(* IEC 61131-3 sources: volt/packages/volt-lsp-iec/test-corpus/twincat-project14/TwinCAT Project14/PLC/Untitled2/Untitled2 Project/References/Tc2_System, 164 files *)

(* ---- E_AdsErr.dut ---- *)
TYPE E_AdsErr :
(
	NOERR,
	ROUTER_NOLOCKEDMEMORY,
	ROUTER_RESIZEMEMORY,
	ROUTER_MAILBOXFULL,
	ROUTER_DEBUGBOXFULL,
	ROUTER_UNKNOWNPORTTYPE,
	ROUTER_NOTINITIALIZED,
	ROUTER_PORTALREADYINUSE,
	ROUTER_NOTREGISTERED,
	ROUTER_NOMOREQUEUES,
	ROUTER_INVALIDPORT,
	ROUTER_NOTACTIVATED,
	ROUTER_FRAGMENTBOXFULL,
	ROUTER_FRAGMENTTIMEOUT,
	ROUTER_TOBEREMOVED,
	DEVICE_ERROR,
	DEVICE_SRVNOTSUPP,
	DEVICE_INVALIDGRP,
	DEVICE_INVALIDOFFSET,
	DEVICE_INVALIDACCESS,
	DEVICE_INVALIDSIZE,
	DEVICE_INVALIDDATA,
	DEVICE_NOTREADY,
	DEVICE_BUSY,
	DEVICE_INVALIDCONTEXT,
	DEVICE_NOMEMORY,
	DEVICE_INVALIDPARM,
	DEVICE_NOTFOUND,
	DEVICE_SYNTAX,
	DEVICE_INCOMPATIBLE,
	DEVICE_EXISTS,
	DEVICE_SYMBOLNOTFOUND,
	DEVICE_SYMBOLVERSIONINVALID,
	DEVICE_INVALIDSTATE,
	DEVICE_TRANSMODENOTSUPP,
	DEVICE_NOTIFYHNDINVALID,
	DEVICE_CLIENTUNKNOWN,
	DEVICE_NOMOREHDLS,
	DEVICE_INVALIDWATCHSIZE,
	DEVICE_NOTINIT,
	DEVICE_TIMEOUT,
	DEVICE_NOINTERFACE,
	DEVICE_INVALIDINTERFACE,
	DEVICE_INVALIDCLSID,
	DEVICE_INVALIDOBJID,
	DEVICE_PENDING,
	DEVICE_ABORTED,
	DEVICE_WARNING,
	DEVICE_INVALIDARRAYIDX,
	DEVICE_SYMBOLNOTACTIVE,
	DEVICE_ACCESSDENIED,
	DEVICE_LICENSENOTFOUND,
	DEVICE_LICENSEEXPIRED,
	DEVICE_LICENSEEXCEEDED,
	DEVICE_LICENSEINVALID,
	DEVICE_LICENSESYSTEMID,
	DEVICE_LICENSENOTIMELIMIT,
	DEVICE_LICENSEFUTUREISSUE,
	DEVICE_LICENSETIMETOLONG,
	DEVICE_EXCEPTION,
	DEVICE_LICENSEDUPLICATED,
	CLIENT_ERROR,
	CLIENT_INVALIDPARM,
	CLIENT_LISTEMPTY,
	CLIENT_VARUSED,
	CLIENT_DUPLINVOKEID,
	CLIENT_SYNCTIMEOUT,
	CLIENT_W32ERROR,
	CLIENT_TIMEOUTINVALID,
	CLIENT_PORTNOTOPEN,
	CLIENT_NOAMSADDR,
	CLIENT_SYNCINTERNAL,
	CLIENT_ADDHASH,
	CLIENT_REMOVEHASH,
	CLIENT_NOMORESYM,
	CLIENT_SYNCRESINVALID,
	CLIENT_SYNCPORTLOCKED
);
END_TYPE

(* ---- E_HRESULTAdsErr.dut ---- *)
TYPE E_HRESULTAdsErr :
(
	HRESULT_ADS_NOERROR,
	ROUTER_NOLOCKEDMEMORY,
	ROUTER_RESIZEMEMORY,
	ROUTER_MAILBOXFULL,
	ROUTER_DEBUGBOXFULL,
	ROUTER_UNKNOWNPORTTYPE,
	ROUTER_NOTINITIALIZED,
	ROUTER_PORTALREADYINUSE,
	ROUTER_NOTREGISTERED,
	ROUTER_NOMOREQUEUES,
	ROUTER_INVALIDPORT,
	ROUTER_NOTACTIVATED,
	ROUTER_FRAGMENTBOXFULL,
	ROUTER_FRAGMENTTIMEOUT,
	ROUTER_TOBEREMOVED,
	ERROR,
	SRVNOTSUPP,
	INVALIDGRP,
	INVALIDOFFSET,
	INVALIDACCESS,
	INVALIDSIZE,
	INVALIDDATA,
	NOTREADY,
	BUSY,
	INVALIDCONTEXT,
	NOMEMORY,
	INVALIDPARM,
	NOTFOUND,
	SYNTAX,
	INCOMPATIBLE,
	EXISTS,
	SYMBOLNOTFOUND,
	SYMBOLVERSIONINVALID,
	INVALIDSTATE,
	TRANSMODENOTSUPP,
	NOTIFYHNDINVALID,
	CLIENTUNKNOWN,
	NOMOREHDLS,
	INVALIDWATCHSIZE,
	NOTINIT,
	TIMEOUT,
	NOINTERFACE,
	INVALIDINTERFACE,
	INVALIDCLSID,
	INVALIDOBJID,
	PENDING,
	ABORTED,
	WARNING,
	INVALIDARRAYIDX,
	SYMBOLNOTACTIVE,
	ACCESSDENIED,
	LICENSENOTFOUND,
	LICENSEEXPIRED,
	LICENSEEXCEEDED,
	LICENSEINVALID,
	LICENSESYSTEMID,
	LICENSENOTIMELIMIT,
	LICENSEFUTUREISSUE,
	LICENSETIMETOLONG,
	EXCEPTION,
	LICENSEDUPLICATED,
	CLIENT_ERROR,
	CLIENT_INVALIDPARM,
	CLIENT_LISTEMPTY,
	CLIENT_VARUSED,
	CLIENT_DUPLINVOKEID,
	CLIENT_SYNCTIMEOUT,
	CLIENT_W32ERROR,
	CLIENT_TIMEOUTINVALID,
	CLIENT_PORTNOTOPEN,
	CLIENT_NOAMSADDR,
	CLIENT_SYNCINTERNAL,
	CLIENT_ADDHASH,
	CLIENT_REMOVEHASH,
	CLIENT_NOMORESYM,
	CLIENT_SYNCRESINVALID,
	CLIENT_SYNCPORTLOCKED
);
END_TYPE

(* ---- E_OpenPath.dut ---- *)
TYPE E_OpenPath :
(
	PATH_GENERIC,
	PATH_BOOTPRJ,
	PATH_BOOTDATA,
	PATH_BOOTPATH,
	PATH_USERPATH1,
	PATH_USERPATH2,
	PATH_USERPATH3,
	PATH_USERPATH4,
	PATH_USERPATH5,
	PATH_USERPATH6,
	PATH_USERPATH7,
	PATH_USERPATH8,
	PATH_USERPATH9
);
END_TYPE

(* ---- E_SeekOrigin.dut ---- *)
TYPE E_SeekOrigin :
(
	SEEK_SET,
	SEEK_CUR,
	SEEK_END
);
END_TYPE

(* ---- E_TcEventClass.dut ---- *)
TYPE E_TcEventClass :
(
	TCEVENTCLASS_NONE,
	TCEVENTCLASS_MAINTENANCE,
	TCEVENTCLASS_MESSAGE,
	TCEVENTCLASS_HINT,
	TCEVENTCLASS_STATEINFO,
	TCEVENTCLASS_INSTRUCTION,
	TCEVENTCLASS_WARNING,
	TCEVENTCLASS_ALARM,
	TCEVENTCLASS_PARAMERROR
);
END_TYPE

(* ---- E_TcEventClearModes.dut ---- *)
TYPE E_TcEventClearModes :
(
	TCEVENTLOGIOFFS_CLEARACTIVE,
	TCEVENTLOGIOFFS_CLEARLOGGED,
	TCEVENTLOGIOFFS_CLEARALL
);
END_TYPE

(* ---- E_TcEventPriority.dut ---- *)
TYPE E_TcEventPriority :
(
	TCEVENTPRIO_IMPLICIT
);
END_TYPE

(* ---- E_TcEventStreamType.dut ---- *)
TYPE E_TcEventStreamType :
(
	TCEVENTSTREAM_INVALID,
	TCEVENTSTREAM_SIMPLE,
	TCEVENTSTREAM_NORMAL,
	TCEVENTSTREAM_NOSOURCE,
	TCEVENTSTREAM_CLASSID,
	TCEVENTSTREAM_CLSNOSRC,
	TCEVENTSTREAM_READCLASSCOUNT,
	TCEVENTSTREAM_MAXTYPE
);
END_TYPE

(* ---- E_TcMemoryArea.dut ---- *)
TYPE E_TcMemoryArea :
(
	Unknown,
	Static,
	Dynamic,
	CNC
);
END_TYPE

(* ---- E_UsrLED_Color.dut ---- *)
TYPE E_UsrLED_Color :
(
	eUsrLED_Off,
	eUsrLED_Red,
	eUsrLED_Blue,
	eUsrLED_Green
);
END_TYPE

(* ---- E_WATCHDOG_TIME_CONFIG.dut ---- *)
TYPE E_WATCHDOG_TIME_CONFIG :
(
	eWATCHDOG_TIME_DISABLED,
	eWATCHDOG_TIME_SECONDS,
	eWATCHDOG_TIME_MINUTES
);
END_TYPE

(* ---- FW_NoOfByte.dut ---- *)
TYPE FW_NoOfByte :
(
	NoOfByte_Byte,
	NoOfByte_Word,
	NoOfByte_DWord
);
END_TYPE

(* ---- Global_Variables.gvl ---- *)
VAR_GLOBAL
	AMSPORT_LOGGER : UINT;
	AMSPORT_EVENTLOG : UINT;
	AMSPORT_R0_RTIME : UINT;
	AMSPORT_R0_IO : UINT;
	AMSPORT_R0_NC : UINT;
	AMSPORT_R0_NCSAF : UINT;
	AMSPORT_R0_NCSVB : UINT;
	AMSPORT_R0_ISG : UINT;
	AMSPORT_R0_CNC : UINT;
	AMSPORT_R0_LINE : UINT;
	AMSPORT_R0_PLC : UINT;
	AMSPORT_R0_PLC_RTS1 : UINT;
	AMSPORT_R0_PLC_RTS2 : UINT;
	AMSPORT_R0_PLC_RTS3 : UINT;
	AMSPORT_R0_PLC_RTS4 : UINT;
	AMSPORT_R0_CAM : UINT;
	AMSPORT_R0_CAMTOOL : UINT;
	AMSPORT_R3_SYSSERV : UINT;
	AMSPORT_R3_SCOPESERVER : UINT;
	ADSSTATE_INVALID : UINT;
	ADSSTATE_IDLE : UINT;
	ADSSTATE_RESET : UINT;
	ADSSTATE_INIT : UINT;
	ADSSTATE_START : UINT;
	ADSSTATE_RUN : UINT;
	ADSSTATE_STOP : UINT;
	ADSSTATE_SAVECFG : UINT;
	ADSSTATE_LOADCFG : UINT;
	ADSSTATE_POWERFAILURE : UINT;
	ADSSTATE_POWERGOOD : UINT;
	ADSSTATE_ERROR : UINT;
	ADSSTATE_SHUTDOWN : UINT;
	ADSSTATE_SUSPEND : UINT;
	ADSSTATE_RESUME : UINT;
	ADSSTATE_CONFIG : UINT;
	ADSSTATE_RECONFIG : UINT;
	ADSSTATE_STOPPING : UINT;
	ADSSTATE_INCOMPATIBLE : UINT;
	ADSSTATE_EXCEPTION : UINT;
	ADSSTATE_MAXSTATES : UINT;
	ADSIGRP_SYMTAB : UDINT;
	ADSIGRP_SYMNAME : UDINT;
	ADSIGRP_SYMVAL : UDINT;
	ADSIGRP_SYM_HNDBYNAME : UDINT;
	ADSIGRP_SYM_VALBYNAME : UDINT;
	ADSIGRP_SYM_VALBYHND : UDINT;
	ADSIGRP_SYM_RELEASEHND : UDINT;
	ADSIGRP_SYM_INFOBYNAME : UDINT;
	ADSIGRP_SYM_VERSION : UDINT;
	ADSIGRP_SYM_INFOBYNAMEEX : UDINT;
	ADSIGRP_SYM_DOWNLOAD : UDINT;
	ADSIGRP_SYM_UPLOAD : UDINT;
	ADSIGRP_SYM_UPLOADINFO : UDINT;
	ADSIGRP_SYMNOTE : UDINT;
	ADSIGRP_IOIMAGE_RWIB : UDINT;
	ADSIGRP_IOIMAGE_RWIX : UDINT;
	ADSIGRP_IOIMAGE_RISIZE : UDINT;
	ADSIGRP_IOIMAGE_RWOB : UDINT;
	ADSIGRP_IOIMAGE_RWOX : UDINT;
	ADSIGRP_IOIMAGE_ROSIZE : UDINT;
	ADSIGRP_IOIMAGE_CLEARI : UDINT;
	ADSIGRP_IOIMAGE_CLEARO : UDINT;
	ADSIGRP_IOIMAGE_RWIOB : UDINT;
	ADSIGRP_DEVICE_DATA : UDINT;
	ADSIOFFS_DEVDATA_ADSSTATE : UDINT;
	ADSIOFFS_DEVDATA_DEVSTATE : UDINT;
	SYSTEMSERVICE_OPENCREATE : UDINT;
	SYSTEMSERVICE_OPENREAD : UDINT;
	SYSTEMSERVICE_OPENWRITE : UDINT;
	SYSTEMSERVICE_CREATEFILE : UDINT;
	SYSTEMSERVICE_CLOSEHANDLE : UDINT;
	SYSTEMSERVICE_FOPEN : UDINT;
	SYSTEMSERVICE_FCLOSE : UDINT;
	SYSTEMSERVICE_FREAD : UDINT;
	SYSTEMSERVICE_FWRITE : UDINT;
	SYSTEMSERVICE_FSEEK : UDINT;
	SYSTEMSERVICE_FTELL : UDINT;
	SYSTEMSERVICE_FGETS : UDINT;
	SYSTEMSERVICE_FPUTS : UDINT;
	SYSTEMSERVICE_FSCANF : UDINT;
	SYSTEMSERVICE_FPRINTF : UDINT;
	SYSTEMSERVICE_FEOF : UDINT;
	SYSTEMSERVICE_FDELETE : UDINT;
	SYSTEMSERVICE_FRENAME : UDINT;
	SYSTEMSERVICE_MKDIR : UDINT;
	SYSTEMSERVICE_RMDIR : UDINT;
	SYSTEMSERVICE_REG_HKEYLOCALMACHINE : UDINT;
	SYSTEMSERVICE_SENDEMAIL : UDINT;
	SYSTEMSERVICE_TIMESERVICES : UDINT;
	SYSTEMSERVICE_STARTPROCESS : UDINT;
	SYSTEMSERVICE_CHANGENETID : UDINT;
	TIMESERVICE_DATEANDTIME : UDINT;
	TIMESERVICE_SYSTEMTIMES : UDINT;
	TIMESERVICE_RTCTIMEDIFF : UDINT;
	TIMESERVICE_ADJUSTTIMETORTC : UDINT;
	TIMESERVICE_TIMEZONINFORMATION : UDINT;
	ADSLOG_MSGTYPE_HINT : DWORD;
	ADSLOG_MSGTYPE_WARN : DWORD;
	ADSLOG_MSGTYPE_ERROR : DWORD;
	ADSLOG_MSGTYPE_LOG : DWORD;
	ADSLOG_MSGTYPE_MSGBOX : DWORD;
	ADSLOG_MSGTYPE_RESOURCE : DWORD;
	ADSLOG_MSGTYPE_STRING : DWORD;
	BOOTDATAFLAGS_RETAIN_LOADED : BYTE;
	BOOTDATAFLAGS_RETAIN_INVALID : BYTE;
	BOOTDATAFLAGS_RETAIN_REQUESTED : BYTE;
	BOOTDATAFLAGS_PERSISTENT_LOADED : BYTE;
	BOOTDATAFLAGS_PERSISTENT_INVALID : BYTE;
	SYSTEMSTATEFLAGS_BSOD : BYTE;
	SYSTEMSTATEFLAGS_RTVIOLATION : BYTE;
	FOPEN_MODEREAD : DWORD;
	FOPEN_MODEWRITE : DWORD;
	FOPEN_MODEAPPEND : DWORD;
	FOPEN_MODEPLUS : DWORD;
	FOPEN_MODEBINARY : DWORD;
	FOPEN_MODETEXT : DWORD;
	FILE_OPENCREATE : DWORD;
	FILE_OPENREAD : DWORD;
	FILE_OPENWRITE : DWORD;
	FILE_READ : DWORD;
	FILE_WRITE : DWORD;
	FILE_SEEKBEGIN : DWORD;
	FILE_SEEKEND : DWORD;
	TCEVENTFLAG_PRIOCLASS : WORD;
	TCEVENTFLAG_FMTSELF : WORD;
	TCEVENTFLAG_LOG : WORD;
	TCEVENTFLAG_MSGBOX : WORD;
	TCEVENTFLAG_SRCID : WORD;
	TCEVENTFLAG_AUTOFMTALL : WORD;
	TCEVENTSTATE_INVALID : WORD;
	TCEVENTSTATE_SIGNALED : WORD;
	TCEVENTSTATE_RESET : WORD;
	TCEVENTSTATE_CONFIRMED : WORD;
	TCEVENTSTATE_RESETCON : WORD;
	TCEVENT_SRCNAMESIZE : INT;
	TCEVENT_FMTPRGSIZE : INT;
	PI : LREAL;
	DEFAULT_ADS_TIMEOUT : TIME;
	MAX_STRING_LENGTH : UDINT;
	MAX_TCBADEV_USERDATA : UDINT;
	SYSTEMSERVICE_BADEVAPI : UDINT;
	BADEVAPIIGRP_GENERAL : UDINT;
	BADEVAPIIOFFS_GENERAL_VERSION : UDINT;
	BIOSIGRP_WATCHDOG : UDINT;
	BIOSIOFFS_WATCHDOG_ENABLE : UDINT;
	BIOSIOFFS_WATCHDOG_CONFIG : UDINT;
	BIOSIOFFS_WATCHDOG_GET_WD_CONFIG : UDINT;
	BIOSIOFFS_WATCHDOG_SET_WD_CONFIG : UDINT;
	BIOSIOFFS_WATCHDOG_ACTIVATE_PWCTR_IO : UDINT;
	BIOSIOFFS_WATCHDOG_TRIG_WD_TIMESPAN : UDINT;
	BIOSIOFFS_WATCHDOG_IO_RETRIGGER : UDINT;
	BIOSIOFFS_WATCHDOG_GET_IO_ADDR : UDINT;
	BIOSIOFFS_WATCHDOG_GET_IO_ADDR_EX : UDINT;
	BIOSIGRP_LED : UDINT;
	BIOSIOFFS_LED_SET_USER : UDINT;
	BIOSIOFFS_LED_SET_USER2 : UDINT;
END_VAR

(* ---- Global_Version.gvl ---- *)
VAR_GLOBAL
	stLibVersion_Tc2_System : ST_LibVersion;
END_VAR

(* ---- Param.gvl ---- *)
VAR_GLOBAL
	TABLE_UPPER_BOUND : INT;
	STRING_LENGTH_EXP : INT;
	STRING_LENGTH_ADDRESS : INT;
	STRING_LENGTH_COMMENT : INT;
	STRING_LENGTH_OUTSTRING : INT;
	TABLE_SHOW_VALID_ITEMS : BOOL;
END_VAR

(* ---- AdsErr_TO_HRESULTAdsErr.pou ---- *)
FUNCTION AdsErr_TO_HRESULTAdsErr : E_HRESULTAdsErr
VAR_INPUT
	eErrId : E_AdsErr;
END_VAR
END_FUNCTION

(* ---- ADSLOGDINT.pou ---- *)
FUNCTION ADSLOGDINT : DINT
VAR_INPUT
	msgCtrlMask : DWORD;
	msgFmtStr : T_MaxString;
	dintArg : DINT;
END_VAR
END_FUNCTION

(* ---- ADSLOGLREAL.pou ---- *)
FUNCTION ADSLOGLREAL : DINT
VAR_INPUT
	msgCtrlMask : DWORD;
	msgFmtStr : T_MaxString;
	lrealArg : LREAL;
END_VAR
END_FUNCTION

(* ---- ADSLOGSTR.pou ---- *)
FUNCTION ADSLOGSTR : DINT
VAR_INPUT
	msgCtrlMask : DWORD;
	msgFmtStr : T_MaxString;
	strArg : T_MaxString;
END_VAR
END_FUNCTION

(* ---- AppendErrorString.pou ---- *)
FUNCTION AppendErrorString
VAR_IN_OUT
	strOld : STRING(STRING_LENGTH_EXP);
	strNew : STRING(1);
END_VAR
END_FUNCTION

(* ---- BAVERSION_TO_DWORD.pou ---- *)
FUNCTION BAVERSION_TO_DWORD : DWORD
VAR_INPUT
	nVersion : BYTE;
	nRevision : BYTE;
	nBuild : WORD;
END_VAR
END_FUNCTION

(* ---- CLEARBIT32.pou ---- *)
FUNCTION CLEARBIT32 : DWORD
VAR_INPUT
	inVal32 : DWORD;
	bitNo : SINT;
END_VAR
END_FUNCTION

(* ---- CONCATX.pou ---- *)
FUNCTION CONCATX
VAR_IN_OUT
	STR1 : STRING(STRING_LENGTH_EXP);
	STR2 : STRING(1);
END_VAR
END_FUNCTION

(* ---- CSETBIT32.pou ---- *)
FUNCTION CSETBIT32 : DWORD
VAR_INPUT
	inVal32 : DWORD;
	bitNo : SINT;
	bitVal : BOOL;
END_VAR
END_FUNCTION

(* ---- F_CheckMemoryArea.pou ---- *)
FUNCTION F_CheckMemoryArea : E_TcMemoryArea
VAR_INPUT
	pData : PVOID;
	nSize : UDINT;
END_VAR
END_FUNCTION

(* ---- F_CmpLibVersion.pou ---- *)
FUNCTION F_CmpLibVersion : DINT
VAR_INPUT
	stVersion : ST_LibVersion;
	iMajor : UINT;
	iMinor : UINT;
	iBuild : UINT;
	iRevision : UINT;
END_VAR
END_FUNCTION

(* ---- F_CompareFwVersion.pou ---- *)
FUNCTION F_CompareFwVersion : BOOL
VAR_INPUT
	major : UINT;
	minor : UINT;
	revision : UINT;
	patch : UINT;
END_VAR
END_FUNCTION

(* ---- F_CreateAmsNetId.pou ---- *)
FUNCTION F_CreateAmsNetId : T_AmsNetId
VAR_INPUT
	nIds : T_AmsNetIdArr;
END_VAR
END_FUNCTION

(* ---- F_CreateIPv4Addr.pou ---- *)
FUNCTION F_CreateIPv4Addr : T_IPv4Addr
VAR_INPUT
	nIds : T_IPv4AddrArr;
END_VAR
END_FUNCTION

(* ---- F_CreateMacAddr.pou ---- *)
FUNCTION F_CreateMacAddr : T_MacAddr
VAR_INPUT
	aMacAddr : T_MacAddrArr;
	sSeparator : STRING(1);
	bLoCase : BOOL;
END_VAR
END_FUNCTION

(* ---- F_GetCpuCoreIndex.pou ---- *)
FUNCTION F_GetCpuCoreIndex : DINT
VAR_INPUT
	nTaskIndex : DINT;
END_VAR
END_FUNCTION

(* ---- F_GetCpuCoreInfo.pou ---- *)
FUNCTION F_GetCpuCoreInfo : HRESULT
VAR_INPUT
	nCpuCoreIndex : DINT;
	pInfo : POINTER TO ST_CpuCoreInfo;
END_VAR
END_FUNCTION

(* ---- F_GetMappingPartner.pou ---- *)
FUNCTION F_GetMappingPartner : OTCID
VAR_INPUT
	p : PVOID;
	n : UDINT;
END_VAR
END_FUNCTION

(* ---- F_GetMappingStatus.pou ---- *)
FUNCTION F_GetMappingStatus : EPlcMappingStatus
VAR_INPUT
	p : PVOID;
	n : UDINT;
END_VAR
END_FUNCTION

(* ---- F_GetStructMemberAlignment.pou ---- *)
FUNCTION F_GetStructMemberAlignment : BYTE
END_FUNCTION

(* ---- F_GetSystemTime.pou ---- *)
FUNCTION F_GetSystemTime : ULINT
END_FUNCTION

(* ---- F_GetTaskInfo.pou ---- *)
FUNCTION F_GetTaskInfo : PlcTaskSystemInfo
END_FUNCTION

(* ---- F_GetTaskTime.pou ---- *)
FUNCTION F_GetTaskTime : ULINT
END_FUNCTION

(* ---- F_GetTaskTotalTime.pou ---- *)
FUNCTION F_GetTaskTotalTime : UDINT
VAR_INPUT
	nTaskIndex : DINT;
END_VAR
END_FUNCTION

(* ---- F_GetVersionTcSystem.pou ---- *)
FUNCTION F_GetVersionTcSystem : UINT
VAR_INPUT
	nVersionElement : INT;
END_VAR
END_FUNCTION

(* ---- F_IOPortRead.pou ---- *)
FUNCTION F_IOPortRead : DWORD
VAR_INPUT
	nAddr : UDINT;
	eSize : E_IOAccessSize;
END_VAR
END_FUNCTION

(* ---- F_IOPortWrite.pou ---- *)
FUNCTION F_IOPortWrite : BOOL
VAR_INPUT
	nAddr : UDINT;
	eSize : E_IOAccessSize;
	nValue : DWORD;
END_VAR
END_FUNCTION

(* ---- F_RaiseException.pou ---- *)
FUNCTION F_RaiseException
VAR_INPUT
	exceptionCode : UDINT;
END_VAR
END_FUNCTION

(* ---- F_ScanAmsNetIds.pou ---- *)
FUNCTION F_ScanAmsNetIds : T_AmsNetIdArr
VAR_INPUT
	sNetID : T_AmsNetID;
END_VAR
END_FUNCTION

(* ---- F_ScanIPv4AddrIds.pou ---- *)
FUNCTION F_ScanIPv4AddrIds : T_IPv4AddrArr
VAR_INPUT
	sIPv4 : T_IPv4Addr;
END_VAR
END_FUNCTION

(* ---- F_SplitPathName.pou ---- *)
FUNCTION F_SplitPathName : BOOL
VAR_INPUT
	sPathName : T_MaxString;
END_VAR
VAR_IN_OUT
	sDrive : STRING(3);
	sDir : T_MaxString;
	sFileName : T_MaxString;
	sExt : T_MaxString;
END_VAR
END_FUNCTION

(* ---- F_ToASC.pou ---- *)
FUNCTION F_ToASC : BYTE
VAR_INPUT
	str : STRING;
END_VAR
END_FUNCTION

(* ---- F_ToCHR.pou ---- *)
FUNCTION F_ToCHR : STRING
VAR_INPUT
	c : BYTE;
END_VAR
END_FUNCTION

(* ---- FW_AdsLogDINT.pou ---- *)
FUNCTION FW_AdsLogDINT : DINT
VAR_INPUT
	nCtrlMask : DWORD;
	sMsgFmt : STRING(255);
	nArg : DINT;
END_VAR
END_FUNCTION

(* ---- FW_AdsLogLREAL.pou ---- *)
FUNCTION FW_AdsLogLREAL : DINT
VAR_INPUT
	nCtrlMask : DWORD;
	sMsgFmt : STRING(255);
	fArg : LREAL;
END_VAR
END_FUNCTION

(* ---- FW_AdsLogSTR.pou ---- *)
FUNCTION FW_AdsLogSTR : DINT
VAR_INPUT
	nCtrlMask : DWORD;
	sMsgFmt : STRING(255);
	sArg : STRING(255);
END_VAR
END_FUNCTION

(* ---- FW_GetCpuIndex.pou ---- *)
FUNCTION FW_GetCpuIndex : DINT
VAR_INPUT
	taskIndex : DINT;
END_VAR
END_FUNCTION

(* ---- FW_GetCpuInfo.pou ---- *)
FUNCTION FW_GetCpuInfo : HRESULT
VAR_INPUT
	cpuIndex : DINT;
	pInfo : POINTER TO ST_CpuCoreInfo;
END_VAR
END_FUNCTION

(* ---- FW_GetCurTaskIndexEx.pou ---- *)
FUNCTION FW_GetCurTaskIndexEx : DINT
END_FUNCTION

(* ---- FW_GetMappingPartner.pou ---- *)
FUNCTION FW_GetMappingPartner : OTCID
VAR_INPUT
	p : PVOID;
	n : UDINT;
END_VAR
END_FUNCTION

(* ---- FW_GetMappingStatus.pou ---- *)
FUNCTION FW_GetMappingStatus : EPlcMappingStatus
VAR_INPUT
	p : PVOID;
	n : UDINT;
END_VAR
END_FUNCTION

(* ---- FW_GetTaskTotalTime.pou ---- *)
FUNCTION FW_GetTaskTotalTime : UDINT
VAR_INPUT
	taskIndex : DINT;
END_VAR
END_FUNCTION

(* ---- FW_GetVersionTcBase.pou ---- *)
FUNCTION FW_GetVersionTcBase : UINT
VAR_INPUT
	nVersionElement : INT;
END_VAR
END_FUNCTION

(* ---- FW_LptSignal.pou ---- *)
FUNCTION FW_LptSignal : BOOL
VAR_INPUT
	nPortAddr : UINT;
	nPinNo : UINT;
	bOnOff : BOOL;
END_VAR
END_FUNCTION

(* ---- FW_MemCmp.pou ---- *)
FUNCTION FW_MemCmp : DINT
VAR_INPUT
	pBuf1 : PVOID;
	pBuf2 : PVOID;
	cbLen : UDINT;
END_VAR
END_FUNCTION

(* ---- FW_MemCpy.pou ---- *)
FUNCTION FW_MemCpy : UDINT
VAR_INPUT
	pDest : PVOID;
	pSrc : PVOID;
	cbLen : UDINT;
END_VAR
END_FUNCTION

(* ---- FW_MemMove.pou ---- *)
FUNCTION FW_MemMove : UDINT
VAR_INPUT
	pDest : PVOID;
	pSrc : PVOID;
	cbLen : UDINT;
END_VAR
END_FUNCTION

(* ---- FW_MemSet.pou ---- *)
FUNCTION FW_MemSet : UDINT
VAR_INPUT
	pDest : PVOID;
	nFillByte : USINT;
	cbLen : UDINT;
END_VAR
END_FUNCTION

(* ---- FW_PortRead.pou ---- *)
FUNCTION FW_PortRead : DWORD
VAR_INPUT
	nPortAddr : UDINT;
	eNoOfByte : FW_NoOfByte;
END_VAR
END_FUNCTION

(* ---- FW_PortWrite.pou ---- *)
FUNCTION FW_PortWrite : BOOL
VAR_INPUT
	nPortAddr : UDINT;
	eNoOfByte : FW_NoOfByte;
	nValue : DWORD;
END_VAR
END_FUNCTION

(* ---- FW_RaiseException.pou ---- *)
FUNCTION FW_RaiseException
VAR_INPUT
	exceptionCode : UDINT;
END_VAR
END_FUNCTION

(* ---- GETBIT32.pou ---- *)
FUNCTION GETBIT32 : BOOL
VAR_INPUT
	inVal32 : DWORD;
	bitNo : SINT;
END_VAR
END_FUNCTION

(* ---- GETCURTASKINDEXEX.pou ---- *)
FUNCTION GETCURTASKINDEXEX : DINT
END_FUNCTION

(* ---- HRESULTAdsErr_TO_AdsErr.pou ---- *)
FUNCTION HRESULTAdsErr_TO_AdsErr : E_AdsErr
VAR_INPUT
	hrErrId : E_HRESULTAdsErr;
END_VAR
END_FUNCTION

(* ---- LPTSIGNAL.pou ---- *)
FUNCTION LPTSIGNAL : BOOL
VAR_INPUT
	PortAddr : UINT;
	PinNo : UINT;
	OnOff : BOOL;
END_VAR
END_FUNCTION

(* ---- MEMCMP.pou ---- *)
FUNCTION MEMCMP : DINT
VAR_INPUT
	pBuf1 : PVOID;
	pBuf2 : PVOID;
	n : UDINT;
END_VAR
END_FUNCTION

(* ---- MEMCPY.pou ---- *)
FUNCTION MEMCPY : UDINT
VAR_INPUT
	destAddr : PVOID;
	srcAddr : PVOID;
	n : UDINT;
END_VAR
END_FUNCTION

(* ---- MEMMOVE.pou ---- *)
FUNCTION MEMMOVE : UDINT
VAR_INPUT
	destAddr : PVOID;
	srcAddr : PVOID;
	n : UDINT;
END_VAR
END_FUNCTION

(* ---- MEMSET.pou ---- *)
FUNCTION MEMSET : UDINT
VAR_INPUT
	destAddr : PVOID;
	fillByte : USINT;
	n : UDINT;
END_VAR
END_FUNCTION

(* ---- ROL32.pou ---- *)
FUNCTION ROL32 : DWORD
VAR_INPUT
	inVal32 : DWORD;
	n : SINT;
END_VAR
END_FUNCTION

(* ---- ROR32.pou ---- *)
FUNCTION ROR32 : DWORD
VAR_INPUT
	inVal32 : DWORD;
	n : SINT;
END_VAR
END_FUNCTION

(* ---- SETBIT32.pou ---- *)
FUNCTION SETBIT32 : DWORD
VAR_INPUT
	inVal32 : DWORD;
	bitNo : SINT;
END_VAR
END_FUNCTION

(* ---- SHL32.pou ---- *)
FUNCTION SHL32 : DWORD
VAR_INPUT
	inVal32 : DWORD;
	n : SINT;
END_VAR
END_FUNCTION

(* ---- SHR32.pou ---- *)
FUNCTION SHR32 : DWORD
VAR_INPUT
	inVal32 : DWORD;
	n : SINT;
END_VAR
END_FUNCTION

(* ---- TestAndSet.pou ---- *)
FUNCTION TestAndSet : BOOL
VAR_IN_OUT
	Flag : BOOL;
END_VAR
END_FUNCTION

(* ---- ADSCLEAREVENTS.pou ---- *)
FUNCTION_BLOCK ADSCLEAREVENTS
VAR_INPUT
	NetID : T_AmsNetId;
	bClear : BOOL;
	iMode : UDINT;
	tTimeout : TIME;
END_VAR
VAR_OUTPUT
	bBusy : BOOL;
	bErr : BOOL;
	iErrId : UDINT;
END_VAR
END_FUNCTION_BLOCK

(* ---- ADSLOGEVENT.pou ---- *)
FUNCTION_BLOCK ADSLOGEVENT
VAR_INPUT
	NETID : T_AmsNetId;
	PORT : UINT;
	Event : BOOL;
	EventQuit : BOOL;
	EventConfigData : TcEvent;
	EventDataAddress : PVOID;
	EventDataLength : UDINT;
	FbCleanup : BOOL;
	TMOUT : TIME;
END_VAR
VAR_OUTPUT
	EventState : UDINT;
	Err : BOOL;
	ErrId : UDINT;
	Quit : BOOL;
END_VAR
END_FUNCTION_BLOCK

(* ---- ADSRDDEVINFO.pou ---- *)
FUNCTION_BLOCK ADSRDDEVINFO
VAR_INPUT
	NETID : T_AmsNetId;
	PORT : T_AmsPort;
	RDINFO : BOOL;
	TMOUT : TIME;
END_VAR
VAR_OUTPUT
	BUSY : BOOL;
	ERR : BOOL;
	ERRID : UDINT;
	DEVNAME : STRING(19);
	DEVVER : UDINT;
END_VAR
END_FUNCTION_BLOCK

(* ---- ADSRDSTATE.pou ---- *)
FUNCTION_BLOCK ADSRDSTATE
VAR_INPUT
	NETID : T_AmsNetId;
	PORT : T_AmsPort;
	RDSTATE : BOOL;
	TMOUT : TIME;
END_VAR
VAR_OUTPUT
	BUSY : BOOL;
	ERR : BOOL;
	ERRID : UDINT;
	ADSSTATE : UINT;
	DEVSTATE : UINT;
END_VAR
END_FUNCTION_BLOCK

(* ---- ADSRDWRT.pou ---- *)
FUNCTION_BLOCK ADSRDWRT
VAR_INPUT
	NETID : T_AmsNetId;
	PORT : T_AmsPort;
	IDXGRP : UDINT;
	IDXOFFS : UDINT;
	WRITELEN : UDINT;
	READLEN : UDINT;
	SRCADDR : PVOID;
	DESTADDR : PVOID;
	WRTRD : BOOL;
	TMOUT : TIME;
END_VAR
VAR_OUTPUT
	BUSY : BOOL;
	ERR : BOOL;
	ERRID : UDINT;
END_VAR
END_FUNCTION_BLOCK

(* ---- ADSRDWRTEX.pou ---- *)
FUNCTION_BLOCK ADSRDWRTEX
VAR_INPUT
	NETID : T_AmsNetId;
	PORT : T_AmsPort;
	IDXGRP : UDINT;
	IDXOFFS : UDINT;
	WRITELEN : UDINT;
	READLEN : UDINT;
	SRCADDR : PVOID;
	DESTADDR : PVOID;
	WRTRD : BOOL;
	TMOUT : TIME;
END_VAR
VAR_OUTPUT
	BUSY : BOOL;
	ERR : BOOL;
	ERRID : UDINT;
	COUNT_R : UDINT;
END_VAR
END_FUNCTION_BLOCK

(* ---- ADSRDWRTIND.pou ---- *)
FUNCTION_BLOCK ADSRDWRTIND
VAR_INPUT
	CLEAR : BOOL;
END_VAR
VAR_OUTPUT
	VALID : BOOL;
	NETID : T_AmsNetId;
	PORT : T_AmsPort;
	INVOKEID : UDINT;
	IDXGRP : UDINT;
	IDXOFFS : UDINT;
	RDLENGTH : UDINT;
	WRTLENGTH : UDINT;
	DATAADDR : PVOID;
END_VAR
END_FUNCTION_BLOCK

(* ---- ADSRDWRTINDEX.pou ---- *)
FUNCTION_BLOCK ADSRDWRTINDEX
VAR_INPUT
	CLEAR : BOOL;
	MINIDXGRP : UDINT;
END_VAR
VAR_OUTPUT
	VALID : BOOL;
	NETID : T_AmsNetId;
	PORT : T_AmsPort;
	INVOKEID : UDINT;
	IDXGRP : UDINT;
	IDXOFFS : UDINT;
	RDLENGTH : UDINT;
	WRTLENGTH : UDINT;
	DATAADDR : PVOID;
END_VAR
END_FUNCTION_BLOCK

(* ---- ADSRDWRTRES.pou ---- *)
FUNCTION_BLOCK ADSRDWRTRES
VAR_INPUT
	NETID : T_AmsNetId;
	PORT : T_AmsPort;
	INVOKEID : UDINT;
	RESULT : UDINT;
	LEN : UDINT;
	DATAADDR : PVOID;
	RESPOND : BOOL;
END_VAR
END_FUNCTION_BLOCK

(* ---- ADSREAD.pou ---- *)
FUNCTION_BLOCK ADSREAD
VAR_INPUT
	NETID : T_AmsNetId;
	PORT : T_AmsPort;
	IDXGRP : UDINT;
	IDXOFFS : UDINT;
	LEN : UDINT;
	DESTADDR : PVOID;
	READ : BOOL;
	TMOUT : TIME;
END_VAR
VAR_OUTPUT
	BUSY : BOOL;
	ERR : BOOL;
	ERRID : UDINT;
END_VAR
END_FUNCTION_BLOCK

(* ---- ADSREADEX.pou ---- *)
FUNCTION_BLOCK ADSREADEX
VAR_INPUT
	NETID : T_AmsNetId;
	PORT : T_AmsPort;
	IDXGRP : UDINT;
	IDXOFFS : UDINT;
	LEN : UDINT;
	DESTADDR : PVOID;
	READ : BOOL;
	TMOUT : TIME;
END_VAR
VAR_OUTPUT
	BUSY : BOOL;
	ERR : BOOL;
	ERRID : UDINT;
	COUNT_R : UDINT;
END_VAR
END_FUNCTION_BLOCK

(* ---- ADSREADIND.pou ---- *)
FUNCTION_BLOCK ADSREADIND
VAR_INPUT
	CLEAR : BOOL;
END_VAR
VAR_OUTPUT
	VALID : BOOL;
	NETID : T_AmsNetId;
	PORT : T_AmsPort;
	INVOKEID : UDINT;
	IDXGRP : UDINT;
	IDXOFFS : UDINT;
	LENGTH : UDINT;
END_VAR
END_FUNCTION_BLOCK

(* ---- ADSREADINDEX.pou ---- *)
FUNCTION_BLOCK ADSREADINDEX
VAR_INPUT
	CLEAR : BOOL;
	MINIDXGRP : UDINT;
END_VAR
VAR_OUTPUT
	VALID : BOOL;
	NETID : T_AmsNetId;
	PORT : T_AmsPort;
	INVOKEID : UDINT;
	IDXGRP : UDINT;
	IDXOFFS : UDINT;
	LENGTH : UDINT;
END_VAR
END_FUNCTION_BLOCK

(* ---- ADSREADRES.pou ---- *)
FUNCTION_BLOCK ADSREADRES
VAR_INPUT
	NETID : T_AmsNetId;
	PORT : T_AmsPort;
	INVOKEID : UDINT;
	RESULT : UDINT;
	LEN : UDINT;
	DATAADDR : PVOID;
	RESPOND : BOOL;
END_VAR
END_FUNCTION_BLOCK

(* ---- ADSWRITE.pou ---- *)
FUNCTION_BLOCK ADSWRITE
VAR_INPUT
	NETID : T_AmsNetId;
	PORT : T_AmsPort;
	IDXGRP : UDINT;
	IDXOFFS : UDINT;
	LEN : UDINT;
	SRCADDR : PVOID;
	WRITE : BOOL;
	TMOUT : TIME;
END_VAR
VAR_OUTPUT
	BUSY : BOOL;
	ERR : BOOL;
	ERRID : UDINT;
END_VAR
END_FUNCTION_BLOCK

(* ---- ADSWRITEIND.pou ---- *)
FUNCTION_BLOCK ADSWRITEIND
VAR_INPUT
	CLEAR : BOOL;
END_VAR
VAR_OUTPUT
	VALID : BOOL;
	NETID : T_AmsNetId;
	PORT : T_AmsPort;
	INVOKEID : UDINT;
	IDXGRP : UDINT;
	IDXOFFS : UDINT;
	LENGTH : UDINT;
	DATAADDR : PVOID;
END_VAR
END_FUNCTION_BLOCK

(* ---- ADSWRITEINDEX.pou ---- *)
FUNCTION_BLOCK ADSWRITEINDEX
VAR_INPUT
	CLEAR : BOOL;
	MINIDXGRP : UDINT;
END_VAR
VAR_OUTPUT
	VALID : BOOL;
	NETID : T_AmsNetId;
	PORT : T_AmsPort;
	INVOKEID : UDINT;
	IDXGRP : UDINT;
	IDXOFFS : UDINT;
	LENGTH : UDINT;
	DATAADDR : PVOID;
END_VAR
END_FUNCTION_BLOCK

(* ---- ADSWRITERES.pou ---- *)
FUNCTION_BLOCK ADSWRITERES
VAR_INPUT
	NETID : T_AmsNetId;
	PORT : T_AmsPort;
	INVOKEID : UDINT;
	RESULT : UDINT;
	RESPOND : BOOL;
END_VAR
END_FUNCTION_BLOCK

(* ---- ADSWRTCTL.pou ---- *)
FUNCTION_BLOCK ADSWRTCTL
VAR_INPUT
	NETID : T_AmsNetId;
	PORT : T_AmsPort;
	ADSSTATE : UINT;
	DEVSTATE : UINT;
	LEN : UDINT;
	SRCADDR : PVOID;
	WRITE : BOOL;
	TMOUT : TIME;
END_VAR
VAR_OUTPUT
	BUSY : BOOL;
	ERR : BOOL;
	ERRID : UDINT;
END_VAR
END_FUNCTION_BLOCK

(* ---- AnalyzeExpression.pou ---- *)
FUNCTION_BLOCK AnalyzeExpression
VAR_INPUT
	InputExp : BOOL;
	DoAnalyze : BOOL;
END_VAR
VAR_OUTPUT
	ExpResult : BOOL;
	OutString : STRING(STRING_LENGTH_OUTSTRING);
END_VAR
END_FUNCTION_BLOCK

(* ---- AnalyzeExpressionCombined.pou ---- *)
FUNCTION_BLOCK AnalyzeExpressionCombined
VAR_INPUT
	InputExp : BOOL;
	DoAnalyze : BOOL;
END_VAR
VAR_OUTPUT
	ExpResult : BOOL;
	OutTable : ARRAY [0..TABLE_UPPER_BOUND] OF ExpressionResult;
	OutString : STRING(STRING_LENGTH_OUTSTRING);
END_VAR
END_FUNCTION_BLOCK

(* ---- AnalyzeExpressionTable.pou ---- *)
FUNCTION_BLOCK AnalyzeExpressionTable
VAR_INPUT
	InputExp : BOOL;
	DoAnalyze : BOOL;
END_VAR
VAR_OUTPUT
	ExpResult : BOOL;
	OutTable : ARRAY [0..TABLE_UPPER_BOUND] OF ExpressionResult;
END_VAR
END_FUNCTION_BLOCK

(* ---- DRAND.pou ---- *)
FUNCTION_BLOCK DRAND
VAR_INPUT
	Seed : INT;
END_VAR
VAR_OUTPUT
	Num : LREAL;
END_VAR
END_FUNCTION_BLOCK

(* ---- FB_AdsReadWriteList.pou ---- *)
FUNCTION_BLOCK FB_AdsReadWriteList
VAR_INPUT
	sNetId : T_AmsNetID;
	nPort : T_AmsPort;
	nIdxGrp : UDINT;
	nIdxOffs : UDINT;
	cbWriteList : UDINT;
	pWriteList : POINTER TO ST_AdsReadWriteListEntry;
	cbReadLen : UDINT;
	pReadBuff : PVOID;
	bExecute : BOOL;
	tTimeout : TIME;
END_VAR
VAR_OUTPUT
	bBusy : BOOL;
	bError : BOOL;
	nErrID : UDINT;
	cbRead : UDINT;
END_VAR
END_FUNCTION_BLOCK

(* ---- FB_BaDeviceIoControl.pou ---- *)
FUNCTION_BLOCK FB_BaDeviceIoControl
VAR_INPUT
	sNetID : T_AmsNetID;
	affinity : T_U64KAFFINITY;
	nModifier : UDINT;
	nIdxGrp : UDINT;
	nIdxOffs : UDINT;
	cbWriteLen : UDINT;
	cbReadLen : UDINT;
	pWriteBuff : PVOID;
	pReadBuff : PVOID;
	bExecute : BOOL;
	tTimeout : TIME;
END_VAR
VAR_OUTPUT
	bBusy : BOOL;
	bError : BOOL;
	nErrID : UDINT;
	cbRead : UDINT;
END_VAR
END_FUNCTION_BLOCK

(* ---- FB_BaGenGetVersion.pou ---- *)
FUNCTION_BLOCK FB_BaGenGetVersion
VAR_INPUT
	sNetID : T_AmsNetID;
	bExecute : BOOL;
	tTimeout : TIME;
END_VAR
VAR_OUTPUT
	bBusy : BOOL;
	bError : BOOL;
	nErrID : UDINT;
	nVersion : BYTE;
	nRevision : BYTE;
	nBuild : WORD;
END_VAR
END_FUNCTION_BLOCK

(* ---- FB_CreateDir.pou ---- *)
FUNCTION_BLOCK FB_CreateDir
VAR_INPUT
	sNetId : T_AmsNetId;
	sPathName : T_MaxString;
	ePath : E_OpenPath;
	bExecute : BOOL;
	tTimeout : TIME;
END_VAR
VAR_OUTPUT
	bBusy : BOOL;
	bError : BOOL;
	nErrId : UDINT;
END_VAR
END_FUNCTION_BLOCK

(* ---- FB_CreateGUID.pou ---- *)
FUNCTION_BLOCK FB_CreateGUID
VAR_INPUT
	bExecute : BOOL;
	sNetId : T_AmsNetId;
	tTimeout : TIME;
	pGuidBuffer : POINTER TO GUID;
	nGuidBufferSize : UDINT;
END_VAR
VAR_OUTPUT
	bBusy : BOOL;
	bError : BOOL;
	nErrorId : UDINT;
END_VAR
END_FUNCTION_BLOCK

(* ---- FB_EOF.pou ---- *)
FUNCTION_BLOCK FB_EOF
VAR_INPUT
	sNetId : T_AmsNetId;
	hFile : UINT;
	bExecute : BOOL;
	tTimeout : TIME;
END_VAR
VAR_OUTPUT
	bBusy : BOOL;
	bError : BOOL;
	nErrId : UDINT;
	bEOF : BOOL;
END_VAR
END_FUNCTION_BLOCK

(* ---- FB_FileClose.pou ---- *)
FUNCTION_BLOCK FB_FileClose
VAR_INPUT
	sNetId : T_AmsNetId;
	hFile : UINT;
	bExecute : BOOL;
	tTimeout : TIME;
END_VAR
VAR_OUTPUT
	bBusy : BOOL;
	bError : BOOL;
	nErrId : UDINT;
END_VAR
END_FUNCTION_BLOCK

(* ---- FB_FileDelete.pou ---- *)
FUNCTION_BLOCK FB_FileDelete
VAR_INPUT
	sNetId : T_AmsNetId;
	sPathName : T_MaxString;
	ePath : E_OpenPath;
	bExecute : BOOL;
	tTimeout : TIME;
END_VAR
VAR_OUTPUT
	bBusy : BOOL;
	bError : BOOL;
	nErrId : UDINT;
END_VAR
END_FUNCTION_BLOCK

(* ---- FB_FileGets.pou ---- *)
FUNCTION_BLOCK FB_FileGets
VAR_INPUT
	sNetId : T_AmsNetId;
	hFile : UINT;
	bExecute : BOOL;
	tTimeout : TIME;
END_VAR
VAR_OUTPUT
	bBusy : BOOL;
	bError : BOOL;
	nErrId : UDINT;
	sLine : T_MaxString;
	bEOF : BOOL;
END_VAR
END_FUNCTION_BLOCK

(* ---- FB_FileLoad.pou ---- *)
FUNCTION_BLOCK FB_FileLoad
VAR_INPUT
	sNetId : T_AmsNetId;
	sPathName : T_MaxString;
	pReadBuff : PVOID;
	cbReadLen : UDINT;
	bExecute : BOOL;
	tTimeout : TIME;
END_VAR
VAR_OUTPUT
	bBusy : BOOL;
	bError : BOOL;
	nErrId : UDINT;
	cbRead : UDINT;
END_VAR
END_FUNCTION_BLOCK

(* ---- FB_FileOpen.pou ---- *)
FUNCTION_BLOCK FB_FileOpen
VAR_INPUT
	sNetId : T_AmsNetId;
	sPathName : T_MaxString;
	nMode : DWORD;
	ePath : E_OpenPath;
	bExecute : BOOL;
	tTimeout : TIME;
END_VAR
VAR_OUTPUT
	bBusy : BOOL;
	bError : BOOL;
	nErrId : UDINT;
	hFile : UINT;
END_VAR
END_FUNCTION_BLOCK

(* ---- FB_FilePuts.pou ---- *)
FUNCTION_BLOCK FB_FilePuts
VAR_INPUT
	sNetId : T_AmsNetId;
	hFile : UINT;
	sLine : T_MaxString;
	bExecute : BOOL;
	tTimeout : TIME;
END_VAR
VAR_OUTPUT
	bBusy : BOOL;
	bError : BOOL;
	nErrId : UDINT;
END_VAR
END_FUNCTION_BLOCK

(* ---- FB_FileRead.pou ---- *)
FUNCTION_BLOCK FB_FileRead
VAR_INPUT
	sNetId : T_AmsNetId;
	hFile : UINT;
	pReadBuff : PVOID;
	cbReadLen : UDINT;
	bExecute : BOOL;
	tTimeout : TIME;
END_VAR
VAR_OUTPUT
	bBusy : BOOL;
	bError : BOOL;
	nErrId : UDINT;
	cbRead : UDINT;
	bEOF : BOOL;
END_VAR
END_FUNCTION_BLOCK

(* ---- FB_FileRename.pou ---- *)
FUNCTION_BLOCK FB_FileRename
VAR_INPUT
	sNetId : T_AmsNetId;
	sOldName : T_MaxString;
	sNewName : T_MaxString;
	ePath : E_OpenPath;
	bExecute : BOOL;
	tTimeout : TIME;
END_VAR
VAR_OUTPUT
	bBusy : BOOL;
	bError : BOOL;
	nErrId : UDINT;
END_VAR
END_FUNCTION_BLOCK

(* ---- FB_FileSeek.pou ---- *)
FUNCTION_BLOCK FB_FileSeek
VAR_INPUT
	sNetId : T_AmsNetId;
	hFile : UINT;
	nSeekPos : DINT;
	eOrigin : E_SeekOrigin;
	bExecute : BOOL;
	tTimeout : TIME;
END_VAR
VAR_OUTPUT
	bBusy : BOOL;
	bError : BOOL;
	nErrId : UDINT;
END_VAR
END_FUNCTION_BLOCK

(* ---- FB_FileTell.pou ---- *)
FUNCTION_BLOCK FB_FileTell
VAR_INPUT
	sNetId : T_AmsNetId;
	hFile : UINT;
	bExecute : BOOL;
	tTimeout : TIME;
END_VAR
VAR_OUTPUT
	bBusy : BOOL;
	bError : BOOL;
	nErrId : UDINT;
	nSeekPos : DINT;
END_VAR
END_FUNCTION_BLOCK

(* ---- FB_FileWrite.pou ---- *)
FUNCTION_BLOCK FB_FileWrite
VAR_INPUT
	sNetId : T_AmsNetId;
	hFile : UINT;
	pWriteBuff : PVOID;
	cbWriteLen : UDINT;
	bExecute : BOOL;
	tTimeout : TIME;
END_VAR
VAR_OUTPUT
	bBusy : BOOL;
	bError : BOOL;
	nErrId : UDINT;
	cbWrite : UDINT;
END_VAR
END_FUNCTION_BLOCK

(* ---- FB_IecCriticalSection.pou ---- *)
FUNCTION_BLOCK FB_IecCriticalSection
END_FUNCTION_BLOCK

(* ---- FB_PcWatchdog.pou ---- *)
FUNCTION_BLOCK FB_PcWatchdog
VAR_INPUT
	tTimeOut : TIME;
	bEnable : BOOL;
END_VAR
VAR_OUTPUT
	bEnabled : BOOL;
	bBusy : BOOL;
	bError : BOOL;
	nErrId : UDINT;
END_VAR
END_FUNCTION_BLOCK

(* ---- FB_PcWatchdog_BAPI.pou ---- *)
FUNCTION_BLOCK FB_PcWatchdog_BAPI
VAR_INPUT
	sNetID : T_AmsNetID;
	nWatchdogTimeS : UDINT (0..15300);
	bExecute : BOOL;
	tTimeout : TIME;
END_VAR
VAR_OUTPUT
	bEnabled : BOOL;
	bBusy : BOOL;
	bError : BOOL;
	nErrID : UDINT;
END_VAR
END_FUNCTION_BLOCK

(* ---- FB_ReadTaskExceedCounter.pou ---- *)
FUNCTION_BLOCK FB_ReadTaskExceedCounter
VAR_INPUT
	bExecute : BOOL;
	nTaskAdsPort : UINT;
END_VAR
VAR_OUTPUT
	bBusy : BOOL;
	bError : BOOL;
	nErrorID : UDINT;
	nExceedCounter : UDINT;
END_VAR
END_FUNCTION_BLOCK

(* ---- FB_RemoveDir.pou ---- *)
FUNCTION_BLOCK FB_RemoveDir
VAR_INPUT
	sNetId : T_AmsNetId;
	sPathName : T_MaxString;
	ePath : E_OpenPath;
	bExecute : BOOL;
	tTimeout : TIME;
END_VAR
VAR_OUTPUT
	bBusy : BOOL;
	bError : BOOL;
	nErrId : UDINT;
END_VAR
END_FUNCTION_BLOCK

(* ---- FB_ResetTaskExceedCounter.pou ---- *)
FUNCTION_BLOCK FB_ResetTaskExceedCounter
VAR_INPUT
	bExecute : BOOL;
	nTaskAdsPort : UINT;
END_VAR
VAR_OUTPUT
	bBusy : BOOL;
	bError : BOOL;
	nErrorID : UDINT;
END_VAR
END_FUNCTION_BLOCK

(* ---- FB_SetLedColor_BAPI.pou ---- *)
FUNCTION_BLOCK FB_SetLedColor_BAPI
VAR_INPUT
	sNetID : T_AmsNetID;
	eNewColor : E_UsrLED_Color;
	bExecute : BOOL;
	tTimeout : TIME;
END_VAR
VAR_OUTPUT
	bBusy : BOOL;
	bError : BOOL;
	nErrID : UDINT;
END_VAR
END_FUNCTION_BLOCK

(* ---- FB_SetLedColorEx_BAPI.pou ---- *)
FUNCTION_BLOCK FB_SetLedColorEx_BAPI
VAR_INPUT
	sNetID : T_AmsNetID;
	nLedID : USINT;
	eNewColor : E_UsrLED_Color;
	bExecute : BOOL;
	tTimeout : TIME;
END_VAR
VAR_OUTPUT
	bBusy : BOOL;
	bError : BOOL;
	nErrID : UDINT;
END_VAR
END_FUNCTION_BLOCK

(* ---- FB_SimpleAdsLogEvent.pou ---- *)
FUNCTION_BLOCK FB_SimpleAdsLogEvent
VAR_INPUT
	SourceID : INT;
	EventID : INT;
	bSetEvent : BOOL;
	bQuit : BOOL;
END_VAR
VAR_OUTPUT
	ErrId : UDINT;
	Error : BOOL;
END_VAR
END_FUNCTION_BLOCK

(* ---- FILECLOSE.pou ---- *)
FUNCTION_BLOCK FILECLOSE
VAR_INPUT
	NETID : T_AmsNetId;
	HFILE : UINT;
	CLOSE : BOOL;
	TMOUT : TIME;
END_VAR
VAR_OUTPUT
	BUSY : BOOL;
	ERR : BOOL;
	ERRID : UDINT;
END_VAR
END_FUNCTION_BLOCK

(* ---- FILEOPEN.pou ---- *)
FUNCTION_BLOCK FILEOPEN
VAR_INPUT
	NETID : T_AmsNetId;
	FPATHNAME : T_MaxString;
	OPENMODE : DWORD;
	OPEN : BOOL;
	TMOUT : TIME;
END_VAR
VAR_OUTPUT
	BUSY : BOOL;
	ERR : BOOL;
	ERRID : UDINT;
	HFILE : UINT;
END_VAR
END_FUNCTION_BLOCK

(* ---- FILEREAD.pou ---- *)
FUNCTION_BLOCK FILEREAD
VAR_INPUT
	NETID : T_AmsNetId;
	HFILE : UINT;
	BUFADDR : PVOID;
	COUNT : UDINT;
	READ : BOOL;
	TMOUT : TIME;
END_VAR
VAR_OUTPUT
	BUSY : BOOL;
	ERR : BOOL;
	ERRID : UDINT;
	COUNT_R : UDINT;
END_VAR
END_FUNCTION_BLOCK

(* ---- FILESEEK.pou ---- *)
FUNCTION_BLOCK FILESEEK
VAR_INPUT
	NETID : T_AmsNetId;
	HFILE : UINT;
	SEEKPOS : UDINT;
	SEEK : BOOL;
	TMOUT : TIME;
END_VAR
VAR_OUTPUT
	BUSY : BOOL;
	ERR : BOOL;
	ERRID : UDINT;
END_VAR
END_FUNCTION_BLOCK

(* ---- FILEWRITE.pou ---- *)
FUNCTION_BLOCK FILEWRITE
VAR_INPUT
	NETID : T_AmsNetId;
	HFILE : UINT;
	BUFADDR : PVOID;
	COUNT : UDINT;
	WRITE : BOOL;
	TMOUT : TIME;
END_VAR
VAR_OUTPUT
	BUSY : BOOL;
	ERR : BOOL;
	ERRID : UDINT;
	COUNT_W : UDINT;
END_VAR
END_FUNCTION_BLOCK

(* ---- FW_AdsClearEvents.pou ---- *)
FUNCTION_BLOCK FW_AdsClearEvents
VAR_INPUT
	sNetId : STRING(23);
	bClear : BOOL;
	nMode : UDINT;
	tTimeout : TIME;
END_VAR
VAR_OUTPUT
	bBusy : BOOL;
	bError : BOOL;
	nErrId : UDINT;
END_VAR
END_FUNCTION_BLOCK

(* ---- FW_AdsLogEvent.pou ---- *)
FUNCTION_BLOCK FW_AdsLogEvent
VAR_INPUT
	sNetId : STRING(23);
	nPort : UINT;
	bEvent : BOOL;
	bEventQuit : BOOL;
	stEventConfigData : FW_TcEvent;
	pEventDataAddress : PVOID;
	cbEventDataLength : UDINT;
	bFbCleanup : BOOL;
	tTimeout : TIME;
END_VAR
VAR_OUTPUT
	nEventState : UDINT;
	bError : BOOL;
	nErrId : UDINT;
	bQuit : BOOL;
END_VAR
END_FUNCTION_BLOCK

(* ---- FW_AdsRdWrt.pou ---- *)
FUNCTION_BLOCK FW_AdsRdWrt
VAR_INPUT
	sNetId : STRING(23);
	nPort : UINT;
	nIdxGrp : UDINT;
	nIdxOffs : UDINT;
	cbWriteLen : UDINT;
	cbReadLen : UDINT;
	pWriteBuff : PVOID;
	pReadBuff : PVOID;
	bExecute : BOOL;
	tTimeout : TIME;
END_VAR
VAR_OUTPUT
	bBusy : BOOL;
	bError : BOOL;
	nErrId : UDINT;
	cbRead : UDINT;
END_VAR
END_FUNCTION_BLOCK

(* ---- FW_AdsRdWrtInd.pou ---- *)
FUNCTION_BLOCK FW_AdsRdWrtInd
VAR_INPUT
	bClear : BOOL;
END_VAR
VAR_OUTPUT
	bValid : BOOL;
	sNetId : STRING(23);
	nPort : UINT;
	nInvokeId : UDINT;
	nIdxGrp : UDINT;
	nIdxOffs : UDINT;
	cbReadLen : UDINT;
	cbWriteLen : UDINT;
	pWriteBuff : PVOID;
END_VAR
END_FUNCTION_BLOCK

(* ---- FW_AdsRdWrtIndEx.pou ---- *)
FUNCTION_BLOCK FW_AdsRdWrtIndEx
VAR_INPUT
	bClear : BOOL;
	nMinIdxGrp : UDINT;
END_VAR
VAR_OUTPUT
	bValid : BOOL;
	sNetId : STRING(23);
	nPort : UINT;
	nInvokeId : UDINT;
	nIdxGrp : UDINT;
	nIdxOffs : UDINT;
	cbReadLen : UDINT;
	cbWriteLen : UDINT;
	pWriteBuff : PVOID;
END_VAR
END_FUNCTION_BLOCK

(* ---- FW_AdsRdWrtList.pou ---- *)
FUNCTION_BLOCK FW_AdsRdWrtList
VAR_INPUT
	sNetId : STRING(23);
	nPort : UINT;
	nIdxGrp : UDINT;
	nIdxOffs : UDINT;
	cbWriteLen : UDINT;
	cbReadLen : UDINT;
	pWriteBuff : POINTER TO ST_AdsReadWriteListEntry;
	pReadBuff : PVOID;
	bExecute : BOOL;
	tTimeout : TIME;
END_VAR
VAR_OUTPUT
	bBusy : BOOL;
	bError : BOOL;
	nErrId : UDINT;
	cbRead : UDINT;
END_VAR
END_FUNCTION_BLOCK

(* ---- FW_AdsRdWrtRes.pou ---- *)
FUNCTION_BLOCK FW_AdsRdWrtRes
VAR_INPUT
	sNetId : STRING(23);
	nPort : UINT;
	nInvokeId : UDINT;
	nErrId : UDINT;
	cbReadLen : UDINT;
	pReadBuff : PVOID;
	bRespond : BOOL;
END_VAR
END_FUNCTION_BLOCK

(* ---- FW_AdsRead.pou ---- *)
FUNCTION_BLOCK FW_AdsRead
VAR_INPUT
	sNetId : STRING(23);
	nPort : UINT;
	nIdxGrp : UDINT;
	nIdxOffs : UDINT;
	cbReadLen : UDINT;
	pReadBuff : PVOID;
	bExecute : BOOL;
	tTimeout : TIME;
END_VAR
VAR_OUTPUT
	bBusy : BOOL;
	bError : BOOL;
	nErrId : UDINT;
	cbRead : UDINT;
END_VAR
END_FUNCTION_BLOCK

(* ---- FW_AdsReadDeviceInfo.pou ---- *)
FUNCTION_BLOCK FW_AdsReadDeviceInfo
VAR_INPUT
	sNetId : STRING(23);
	nPort : UINT;
	bExecute : BOOL;
	tTimeout : TIME;
END_VAR
VAR_OUTPUT
	bBusy : BOOL;
	bError : BOOL;
	nErrId : UDINT;
	sDevName : STRING(19);
	nDevVersion : UDINT;
END_VAR
END_FUNCTION_BLOCK

(* ---- FW_AdsReadInd.pou ---- *)
FUNCTION_BLOCK FW_AdsReadInd
VAR_INPUT
	bClear : BOOL;
END_VAR
VAR_OUTPUT
	bValid : BOOL;
	sNetId : STRING(23);
	nPort : UINT;
	nInvokeId : UDINT;
	nIdxGrp : UDINT;
	nIdxOffs : UDINT;
	cbReadLen : UDINT;
END_VAR
END_FUNCTION_BLOCK

(* ---- FW_AdsReadIndEx.pou ---- *)
FUNCTION_BLOCK FW_AdsReadIndEx
VAR_INPUT
	bClear : BOOL;
	nMinIdxGrp : UDINT;
END_VAR
VAR_OUTPUT
	bValid : BOOL;
	sNetId : STRING(23);
	nPort : UINT;
	nInvokeId : UDINT;
	nIdxGrp : UDINT;
	nIdxOffs : UDINT;
	cbReadLen : UDINT;
END_VAR
END_FUNCTION_BLOCK

(* ---- FW_AdsReadRes.pou ---- *)
FUNCTION_BLOCK FW_AdsReadRes
VAR_INPUT
	sNetId : STRING(23);
	nPort : UINT;
	nInvokeId : UDINT;
	nErrId : UDINT;
	cbReadLen : UDINT;
	pReadBuff : PVOID;
	bRespond : BOOL;
END_VAR
END_FUNCTION_BLOCK

(* ---- FW_AdsReadState.pou ---- *)
FUNCTION_BLOCK FW_AdsReadState
VAR_INPUT
	sNetId : STRING(23);
	nPort : UINT;
	bExecute : BOOL;
	tTimeout : TIME;
END_VAR
VAR_OUTPUT
	bBusy : BOOL;
	bError : BOOL;
	nErrId : UDINT;
	nAdsState : UINT;
	nDevState : UINT;
END_VAR
END_FUNCTION_BLOCK

(* ---- FW_AdsWrite.pou ---- *)
FUNCTION_BLOCK FW_AdsWrite
VAR_INPUT
	sNetId : STRING(23);
	nPort : UINT;
	nIdxGrp : UDINT;
	nIdxOffs : UDINT;
	cbWriteLen : UDINT;
	pWriteBuff : PVOID;
	bExecute : BOOL;
	tTimeout : TIME;
END_VAR
VAR_OUTPUT
	bBusy : BOOL;
	bError : BOOL;
	nErrId : UDINT;
END_VAR
END_FUNCTION_BLOCK

(* ---- FW_AdsWriteControl.pou ---- *)
FUNCTION_BLOCK FW_AdsWriteControl
VAR_INPUT
	sNetId : STRING(23);
	nPort : UINT;
	nAdsState : UINT;
	nDevState : UINT;
	cbWriteLen : UDINT;
	pWriteBuff : PVOID;
	bExecute : BOOL;
	tTimeout : TIME;
END_VAR
VAR_OUTPUT
	bBusy : BOOL;
	bError : BOOL;
	nErrId : UDINT;
END_VAR
END_FUNCTION_BLOCK

(* ---- FW_AdsWriteInd.pou ---- *)
FUNCTION_BLOCK FW_AdsWriteInd
VAR_INPUT
	bClear : BOOL;
END_VAR
VAR_OUTPUT
	bValid : BOOL;
	sNetId : STRING(23);
	nPort : UINT;
	nInvokeId : UDINT;
	nIdxGrp : UDINT;
	nIdxOffs : UDINT;
	cbWriteLen : UDINT;
	pWriteBuff : PVOID;
END_VAR
END_FUNCTION_BLOCK

(* ---- FW_AdsWriteIndEx.pou ---- *)
FUNCTION_BLOCK FW_AdsWriteIndEx
VAR_INPUT
	bClear : BOOL;
	nMinIdxGrp : UDINT;
END_VAR
VAR_OUTPUT
	bValid : BOOL;
	sNetId : STRING(23);
	nPort : UINT;
	nInvokeId : UDINT;
	nIdxGrp : UDINT;
	nIdxOffs : UDINT;
	cbWriteLen : UDINT;
	pWriteBuff : PVOID;
END_VAR
END_FUNCTION_BLOCK

(* ---- FW_AdsWriteRes.pou ---- *)
FUNCTION_BLOCK FW_AdsWriteRes
VAR_INPUT
	sNetId : STRING(23);
	nPort : UINT;
	nInvokeId : UDINT;
	nErrId : UDINT;
	bRespond : BOOL;
END_VAR
END_FUNCTION_BLOCK

(* ---- FW_DRand.pou ---- *)
FUNCTION_BLOCK FW_DRand
VAR_INPUT
	nSeed : INT;
END_VAR
VAR_OUTPUT
	fRndNum : LREAL;
END_VAR
END_FUNCTION_BLOCK

(* ---- FW_GetCpuAccount.pou ---- *)
FUNCTION_BLOCK FW_GetCpuAccount
VAR_OUTPUT
	dwCpuAccount : UDINT;
END_VAR
END_FUNCTION_BLOCK

(* ---- FW_GetCpuCounter.pou ---- *)
FUNCTION_BLOCK FW_GetCpuCounter
VAR_OUTPUT
	dwCpuCntLo : UDINT;
	dwCpuCntHi : UDINT;
END_VAR
END_FUNCTION_BLOCK

(* ---- FW_GetCurTaskIndex.pou ---- *)
FUNCTION_BLOCK FW_GetCurTaskIndex
VAR_OUTPUT
	nIndex : BYTE;
END_VAR
END_FUNCTION_BLOCK

(* ---- FW_GetSystemTime.pou ---- *)
FUNCTION_BLOCK FW_GetSystemTime
VAR_OUTPUT
	dwTimeLo : UDINT;
	dwTimeHi : UDINT;
END_VAR
END_FUNCTION_BLOCK

(* ---- FW_GetTaskTime.pou ---- *)
FUNCTION_BLOCK FW_GetTaskTime
VAR_OUTPUT
	timeLoDW : UDINT;
	timeHiDW : UDINT;
END_VAR
END_FUNCTION_BLOCK

(* ---- GETCPUACCOUNT.pou ---- *)
FUNCTION_BLOCK GETCPUACCOUNT
VAR_OUTPUT
	cpuAccountDW : UDINT;
END_VAR
END_FUNCTION_BLOCK

(* ---- GETCPUCOUNTER.pou ---- *)
FUNCTION_BLOCK GETCPUCOUNTER
VAR_OUTPUT
	cpuCntLoDW : UDINT;
	cpuCntHiDW : UDINT;
END_VAR
END_FUNCTION_BLOCK

(* ---- GETCURTASKINDEX.pou ---- *)
FUNCTION_BLOCK GETCURTASKINDEX
VAR_OUTPUT
	index : BYTE;
END_VAR
END_FUNCTION_BLOCK

(* ---- GETSYSTEMTIME.pou ---- *)
FUNCTION_BLOCK GETSYSTEMTIME
VAR_OUTPUT
	timeLoDW : UDINT;
	timeHiDW : UDINT;
END_VAR
END_FUNCTION_BLOCK

(* ---- GETTASKTIME.pou ---- *)
FUNCTION_BLOCK GETTASKTIME
VAR_OUTPUT
	timeLoDW : UDINT;
	timeHiDW : UDINT;
END_VAR
END_FUNCTION_BLOCK

(* ---- SFCActionControl.pou ---- *)
FUNCTION_BLOCK SFCActionControl
VAR_INPUT
	N : BOOL;
	R0 : BOOL;
	S0 : BOOL;
	L : BOOL;
	D : BOOL;
	P : BOOL;
	SD : BOOL;
	DS : BOOL;
	SL : BOOL;
	T : TIME;
END_VAR
VAR_OUTPUT
	Q : BOOL;
END_VAR
END_FUNCTION_BLOCK
